// TIA Portal V20 export
// export: Created 2026-10-20T18:55:11.8487258Z, ExportSetting None, DisplayName Totally Integrated Automation Portal, DisplayVersion V20 Update 6, DisplayName TIA Portal Openness, DisplayVersion V20 Update 6, DisplayName TIA Portal Version Control Interface, DisplayVersion V20 Update 6, DisplayName SINAMICS Startdrive Advanced, DisplayVersion V20 SP1, DisplayName SINAMICS Startdrive G130, G150, S120, S150, SINAMICS MV, G220, S200, S210, DisplayVersion V20 SP1, DisplayName SINAMICS Startdrive G110M, G120, G120C, G120D, G120P, G115D, DisplayVersion V20 SP1, DisplayName STEP 7 Professional, DisplayVersion V20 Update 6, DisplayName STEP 7 Safety, DisplayVersion V20 Update 2, DisplayName WinCC Basic/Comfort/Advanced, DisplayVersion V20 Update 6, DisplayName WinCC Unified, DisplayVersion V20 Update 6
VAR_GLOBAL   // PLC tag table "IO_VFDs_4"
   C4107_StatusWord AT %IW2702 : Word;
   C4106_ActualSpeed AT %IW2692 : Word;
   C4103_MainSetpoint AT %QW1219 : Word;
   C4101_StatusWord AT %IW2630 : Word;
   C4105_ActualCurrent AT %IW2682 : Word;
   C4102_ActualSpeed AT %IW2644 : Word;
   C4103_ActualSpeed AT %IW2656 : Word;
   C4102_MainSetpoint AT %QW1177 : Word;
   C4104_MainSetpoint AT %QW1223 : Word;
   C4106_ActualCurrent AT %IW2694 : Word;
   C4106_MainSetpoint AT %QW1231 : Word;
   C4107_ControlWord AT %QW1233 : Word;
   VTD4_ActualSpeed AT %IW1331 : Word;
   C4108_ActualCurrent AT %IW2718 : Word;
   CVTD4_ActualCurrent AT %IW2622 : Word;
   CVTD4_MainSetpoint AT %QW1169 : Word;
   CVTD4_ActualSpeed AT %IW2620 : Word;
   C4102_ActualCurrent AT %IW2646 : Word;
   C4105_StatusWord AT %IW2678 : Word;
   C4105_MainSetpoint AT %QW1227 : Word;
   C4101_ActualCurrent AT %IW2634 : Word;
   C4104_StatusWord AT %IW2666 : Word;
   CVTD4_StatusWord AT %IW2618 : Word;
   C4102_ControlWord AT %QW1175 : Word;
   C4108_MainSetpoint AT %QW1239 : Word;
   C4108_ActualSpeed AT %IW2716 : Word;
   C4103_ActualCurrent AT %IW2658 : Word;
   C4104_ActualCurrent AT %IW2670 : Word;
   C4106_StatusWord AT %IW2690 : Word;
   C4101_ActualSpeed AT %IW2632 : Word;
   C4108_ControlWord AT %QW1237 : Word;
   C4104_ActualSpeed AT %IW2668 : Word;
   VTD4_ActualCurrent AT %IW1333 : Word;
   C4101_ControlWord AT %QW1171 : Word;
   VTD4_MainSetpoint AT %QW1165 : Word;
   C4107_ActualCurrent AT %IW2706 : Word;
   VTD4_ControlWord AT %QW1163 : Word;
   C4105_ControlWord AT %QW1225 : Word;
   C4101_MainSetpoint AT %QW1173 : Word;
   C4106_ControlWord AT %QW1229 : Word;
   C4104_ControlWord AT %QW1221 : Word;
   C4103_ControlWord AT %QW1217 : Word;
   VTD4_StatusWord AT %IW1329 : Word;
   C4108_StatusWord AT %IW2714 : Word;
   C4107_MainSetpoint AT %QW1235 : Word;
   C4105_ActualSpeed AT %IW2680 : Word;
   C4103_StatusWord AT %IW2654 : Word;
   C4107_ActualSpeed AT %IW2704 : Word;
   C4102_StatusWord AT %IW2642 : Word;
   CVTD4_ControlWord AT %QW1167 : Word;
   C4104_ActualTorque AT %IW2672 : Word;
   VTD4_ActualTorque AT %IW1336 : Word;
   C4106_ActualTorque AT %IW2696 : Word;
   C4108_ActualTorque AT %IW2720 : Word;
   C4103_ActualTorque AT %IW2660 : Word;
   C4101_ActualTorque AT %IW2636 : Word;
   C4105_ActualTorque AT %IW2684 : Word;
   C4107_ActualTorque AT %IW2708 : Word;
   CVTD4_ActualTorque AT %IW2624 : Word;
   C4102_ActualTorque AT %IW2648 : Word;
   VTD4_AccFactor AT %QW1525 : Word;
END_VAR
